(* Logix 5000 project; controller TFF vendor 1 type 14 code 107 rev 33.11; software revision 33.04; part 34 of 38 *)
(* tags used below, declared in another part *)
   Address : DINT;   // Temp Address
   Index : DINT;   // Index
   Index2 : DINT;   // Index
   _150S1 : ALIAS FOR DigitalOutput[0];
   AC008 : ALIAS FOR DigitalOutput[7];
   AlarmControl : AlarmControl;   // Alarm Control
   ALM001 : ALIAS FOR DigitalOutput[2];
   ALM002 : ALIAS FOR DigitalOutput[17];
   AnalogOutput : AnalogOutput[25];   // Analog Output Array
   AO1 : ALIAS FOR AnalogOutput[8];
   AO2 : ALIAS FOR AnalogOutput[9];
   AO3 : ALIAS FOR AnalogOutput[10];
   AO4 : ALIAS FOR AnalogOutput[11];
   AP008 : ALIAS FOR DigitalOutput[14];
   BAN001P : ALIAS FOR DigitalOutput[4];
   BAN001S : ALIAS FOR DigitalOutput[3];
   BAN002P : ALIAS FOR DigitalOutput[6];
   BAN002S : ALIAS FOR DigitalOutput[5];
   DigitalOutput : BOOL[256];   // Digital Output Array these bits are sent to output cards.
   DO1 : ALIAS FOR DigitalOutput[80];
   DO2 : ALIAS FOR DigitalOutput[81];
   DO3 : ALIAS FOR DigitalOutput[82];
   DO4 : ALIAS FOR DigitalOutput[83];
   DO5 : ALIAS FOR DigitalOutput[84];
   DO6 : ALIAS FOR DigitalOutput[85];
   DO7 : ALIAS FOR DigitalOutput[86];
   FlowPath : FlowPath[64];   // Flow Path Array
   IBA001 : ALIAS FOR DigitalOutput[25];
   MIX101ON : ALIAS FOR DigitalOutput[16];
   Mixer : Mixer;   // Mixer config. structure
   PCV101 : ALIAS FOR AnalogPoint[3];
   PCV101_AO : ALIAS FOR AnalogOutput[3];
   PCV201 : ALIAS FOR AnalogPoint[4];
   PCV201_AO : ALIAS FOR AnalogOutput[4];
   POWERON : ALIAS FOR DigitalOutput[1];
   PTA001 : ALIAS FOR DigitalOutput[21];
   PTA101 : ALIAS FOR DigitalOutput[22];
   PTA201 : ALIAS FOR DigitalOutput[23];
   PTA401 : ALIAS FOR DigitalOutput[24];
   PTA601 : ALIAS FOR DigitalOutput[26];
   Rack_Murr_Node0_Smart : IO_Station;   // Status of Node 0 Smart
   Rack_Murr_Node1_TFF40 : IO_Station;   // Status of Node 1 TFF40
   Rack_Murr_Node1_TFF80 : IO_Station;   // Status of Node 1 TFF80
   SIC001 : ALIAS FOR Drive[1];
   SIC001_AO : ALIAS FOR AnalogOutput[0];
   SIC001_DO : ALIAS FOR DigitalOutput[8];
   SIC002 : ALIAS FOR Drive[2];
   SIC002_AO : ALIAS FOR AnalogOutput[1];
   SIC002_DO : ALIAS FOR DigitalOutput[9];
   SIC003_AO : ALIAS FOR AnalogOutput[2];
   SIC003_DO : ALIAS FOR DigitalOutput[15];
   SIC004 : ALIAS FOR Drive[3];
   SIC004_AO : ALIAS FOR AnalogOutput[5];
   SysControl : SysControl;   // General system status and command
   Tank : TankManagement;   // Tank Management
   TCU101 : ALIAS FOR AnalogPoint[18];
   TCU101_AO : ALIAS FOR AnalogOutput[6];
   TCU101ON : ALIAS FOR DigitalOutput[20];
   ThisSystem : SystemType;
   TNK101 : ALIAS FOR DigitalOutput[18];
   TNK102 : ALIAS FOR DigitalOutput[19];
   TNK103 : ALIAS FOR DigitalOutput[27];
   Valve : Valve[100];   // Valve Array
   ValveControl : ValveControl;   // Valve Control
   XV001 : ALIAS FOR Valve[0];
   XV002 : ALIAS FOR Valve[1];
   XV003 : ALIAS FOR Valve[2];
   XV004 : ALIAS FOR Valve[3];
   XV005 : ALIAS FOR Valve[4];
   XV006 : ALIAS FOR Valve[5];
   XV007 : ALIAS FOR Valve[6];
   XV101 : ALIAS FOR Valve[7];
   XV102 : ALIAS FOR Valve[8];
   XV201 : ALIAS FOR Valve[15];
   XV202 : ALIAS FOR Valve[16];
   XV401 : ALIAS FOR Valve[9];
   XV402 : ALIAS FOR Valve[10];
   XV403 : ALIAS FOR Valve[11];
   XV404 : ALIAS FOR Valve[12];
   XV405 : ALIAS FOR Valve[13];
   XV406 : ALIAS FOR Valve[14];
   XV701 : ALIAS FOR Valve[17];
   XV702 : ALIAS FOR Valve[18];
   XV703 : ALIAS FOR Valve[19];
   XV704 : ALIAS FOR Valve[20];
   Y500A : ALIAS FOR DigitalOutput[10];
   Y500B : ALIAS FOR DigitalOutput[11];
   Y501A : ALIAS FOR DigitalOutput[12];
   Y501B : ALIAS FOR DigitalOutput[13];
(* Process, continued *)

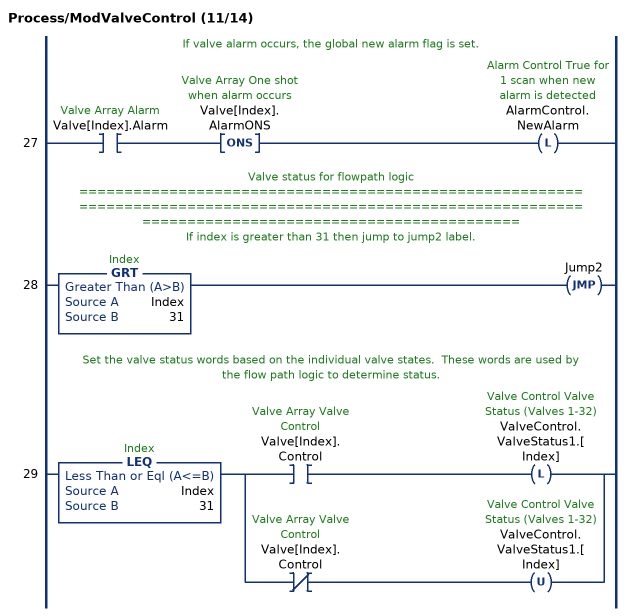
   [picture p422: Process/ModValveControl rungs 27-29]
   // If valve alarm occurs, the global new alarm flag is set.
   27: XIC(Valve[Index].Alarm)ONS(Valve[Index].AlarmONS)OTL(AlarmControl.NewAlarm);
   // Valve status for flowpath logic
   // ==========================================================================================================================================================
   // If index is greater than 31 then jump to jump2 label.
   28: GRT(Index,31)JMP(Jump2);
   // Set the valve status words based on the individual valve states.  These words are used by the flow path logic to determine status.
   29: LEQ(Index,31)[XIC(Valve[Index].Control) OTL(ValveControl.ValveStatus1.[Index]) ,XIO(Valve[Index].Control) OTU(ValveControl.ValveStatus1.[Index]) ];
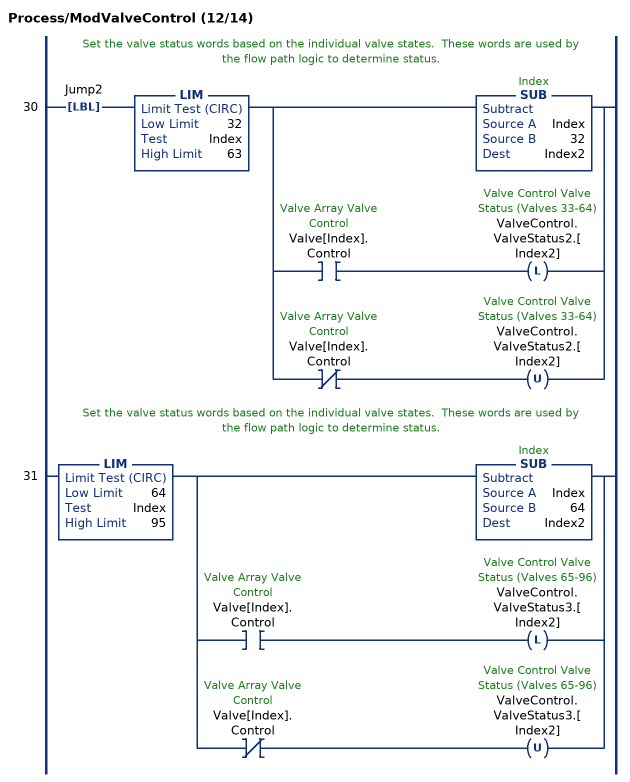
   // Set the valve status words based on the individual valve states.  These words are used by the flow path logic to determine status.
   30: LBL(Jump2)LIM(32,Index,63)[SUB(Index,32,Index2) ,XIC(Valve[Index].Control) OTL(ValveControl.ValveStatus2.[Index2]) ,XIO(Valve[Index].Control) OTU(ValveControl.ValveStatus2.[Index2]) ];
   // Set the valve status words based on the individual valve states.  These words are used by the flow path logic to determine status.
   31: LIM(64,Index,95)[SUB(Index,64,Index2) ,XIC(Valve[Index].Control) OTL(ValveControl.ValveStatus3.[Index2]) ,XIO(Valve[Index].Control) OTU(ValveControl.ValveStatus3.[Index2]) ];
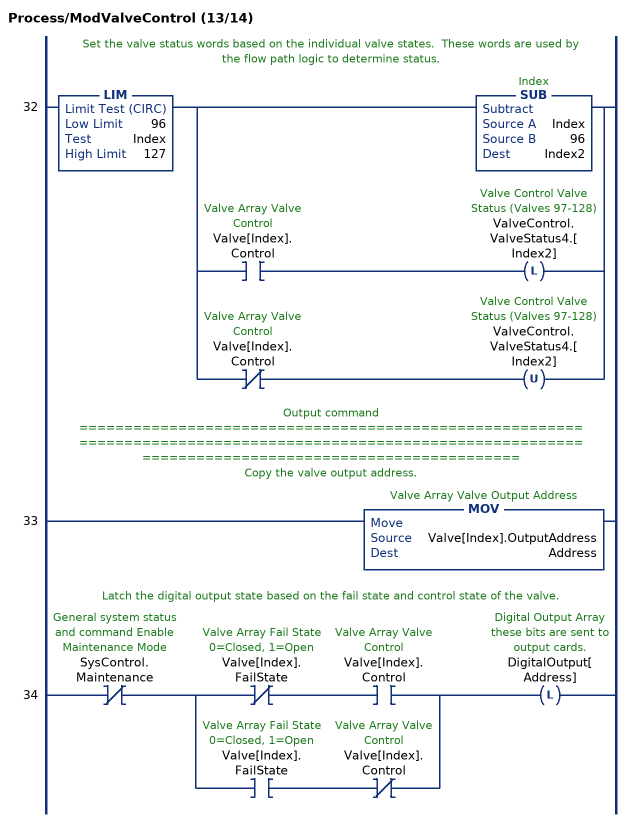
   // Set the valve status words based on the individual valve states.  These words are used by the flow path logic to determine status.
   32: LIM(96,Index,127)[SUB(Index,96,Index2) ,XIC(Valve[Index].Control) OTL(ValveControl.ValveStatus4.[Index2]) ,XIO(Valve[Index].Control) OTU(ValveControl.ValveStatus4.[Index2]) ];
   // Output command
   // ==========================================================================================================================================================
   // Copy the valve output address.
   33: MOV(Valve[Index].OutputAddress,Address);
   // Latch the digital output state based on the fail state and control state of the valve.
   34: XIO(SysControl.Maintenance)[XIO(Valve[Index].FailState) XIC(Valve[Index].Control) ,XIC(Valve[Index].FailState) XIO(Valve[Index].Control) ]OTL(DigitalOutput[Address]);
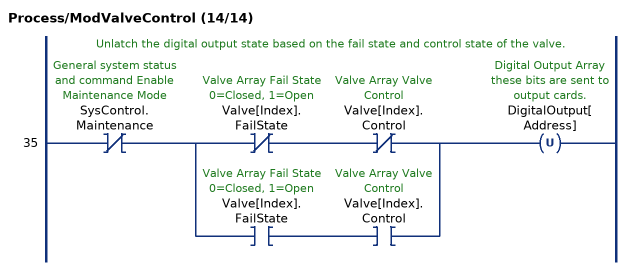
   // Unlatch the digital output state based on the fail state and control state of the valve.
   35: XIO(SysControl.Maintenance)[XIO(Valve[Index].FailState) XIO(Valve[Index].Control) ,XIC(Valve[Index].FailState) XIC(Valve[Index].Control) ]OTU(DigitalOutput[Address]);
END_ROUTINE

ROUTINE OutputAnalogPoint   (* ladder *)
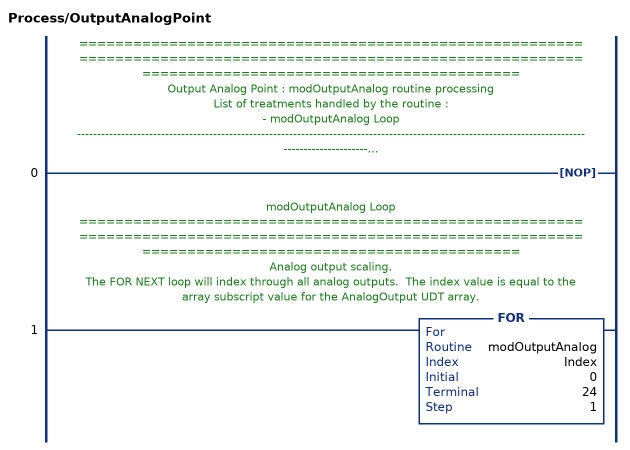
   // ==========================================================================================================================================================
   //                                                                                                             Output Analog Point : modOutputAnalog routine processing
   //                                                     List of treatments handled by the routine :
   //                                                          - modOutputAnalog Loop
   //                                                     -----------------------------------------------------------------------------------------------------------------------------------------------------
   //                                                     History
   // 		2019-DEC-24 - Merck - Q. Spindler - Initial version for Candidate Release 1.00.00.00.a
   // ==========================================================================================================================================================
   0: NOP();
   // modOutputAnalog Loop
   // ==========================================================================================================================================================
   // Analog output scaling.
   // The FOR NEXT loop will index through all analog outputs.  The index value is equal to the array subscript value for the AnalogOutput UDT array.
   1: FOR(modOutputAnalog,Index,0,24,1);
END_ROUTINE

ROUTINE OutputAnalogRaw   (* ladder *)
// Output Routine
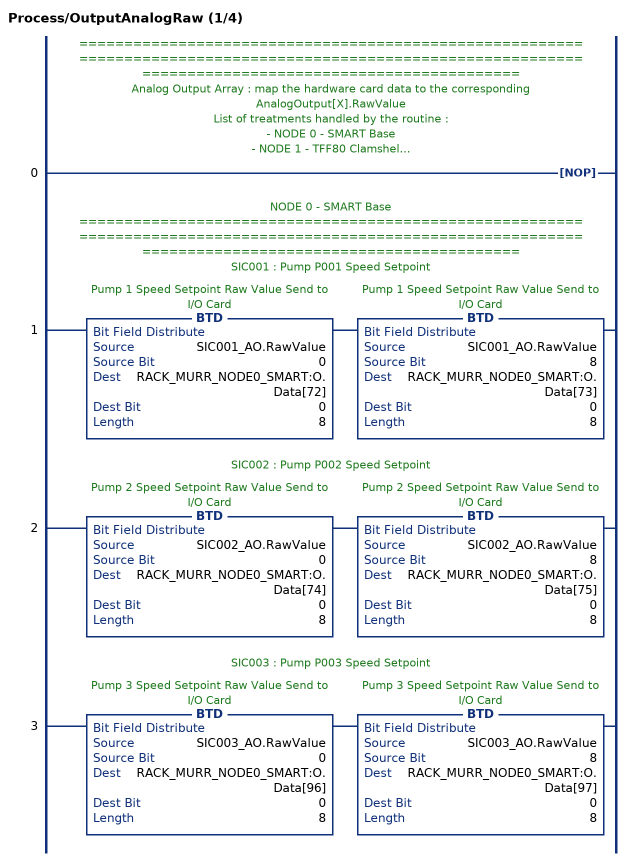
   // ==========================================================================================================================================================
   //                                                                                    Analog Output Array : map the hardware card data to the corresponding AnalogOutput[X].RawValue
   //                                                     List of treatments handled by the routine :
   //                                                    - NODE 0 - SMART Base
   //                                                         - NODE 1 - TFF80 Clamshell
   //                                                         - NODE 1 - TFF40 Clamshell
   //                                                         - NODE 1 - TFF20 Clamshell
   //                                                     -----------------------------------------------------------------------------------------------------------------------------------------------------
   //                                                     History
   // 		2019-DEC-24 - Merck - Q. Spindler - Initial version for Candidate Release 1.00.00.00.a
   // ==========================================================================================================================================================
   0: NOP();
   // NODE 0 - SMART Base
   // ==========================================================================================================================================================
   // SIC001 : Pump P001 Speed Setpoint
   1: BTD(SIC001_AO.RawValue,0,RACK_MURR_NODE0_SMART:O.Data[72],0,8)BTD(SIC001_AO.RawValue,8,RACK_MURR_NODE0_SMART:O.Data[73],0,8);
   // SIC002 : Pump P002 Speed Setpoint
   2: BTD(SIC002_AO.RawValue,0,RACK_MURR_NODE0_SMART:O.Data[74],0,8)BTD(SIC002_AO.RawValue,8,RACK_MURR_NODE0_SMART:O.Data[75],0,8);
   // SIC003 : Pump P003 Speed Setpoint
   3: BTD(SIC003_AO.RawValue,0,RACK_MURR_NODE0_SMART:O.Data[96],0,8)BTD(SIC003_AO.RawValue,8,RACK_MURR_NODE0_SMART:O.Data[97],0,8);
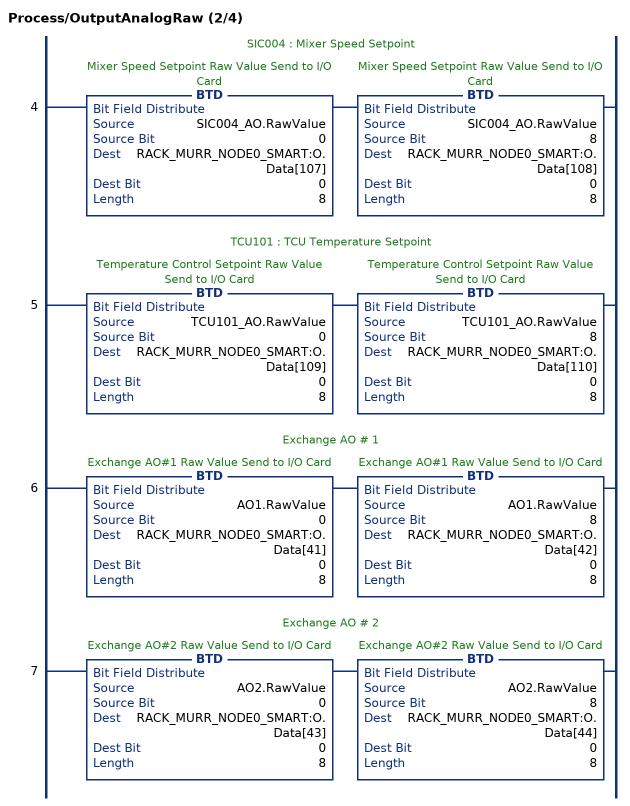
   // SIC004 : Mixer Speed Setpoint
   4: BTD(SIC004_AO.RawValue,0,RACK_MURR_NODE0_SMART:O.Data[107],0,8)BTD(SIC004_AO.RawValue,8,RACK_MURR_NODE0_SMART:O.Data[108],0,8);
   // TCU101 : TCU Temperature Setpoint
   5: BTD(TCU101_AO.RawValue,0,RACK_MURR_NODE0_SMART:O.Data[109],0,8)BTD(TCU101_AO.RawValue,8,RACK_MURR_NODE0_SMART:O.Data[110],0,8);
   // Exchange AO # 1
   6: BTD(AO1.RawValue,0,RACK_MURR_NODE0_SMART:O.Data[41],0,8)BTD(AO1.RawValue,8,RACK_MURR_NODE0_SMART:O.Data[42],0,8);
   // Exchange AO # 2
   7: BTD(AO2.RawValue,0,RACK_MURR_NODE0_SMART:O.Data[43],0,8)BTD(AO2.RawValue,8,RACK_MURR_NODE0_SMART:O.Data[44],0,8);
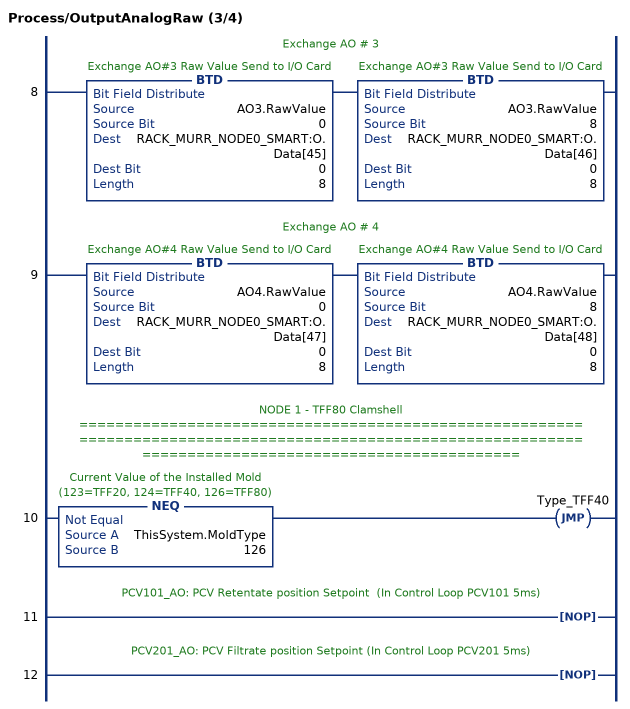
   // Exchange AO # 3
   8: BTD(AO3.RawValue,0,RACK_MURR_NODE0_SMART:O.Data[45],0,8)BTD(AO3.RawValue,8,RACK_MURR_NODE0_SMART:O.Data[46],0,8);
   // Exchange AO # 4
   9: BTD(AO4.RawValue,0,RACK_MURR_NODE0_SMART:O.Data[47],0,8)BTD(AO4.RawValue,8,RACK_MURR_NODE0_SMART:O.Data[48],0,8);
   // NODE 1 - TFF80 Clamshell
   // ==========================================================================================================================================================
   10: NEQ(ThisSystem.MoldType,126)JMP(Type_TFF40);
   // PCV101_AO: PCV Retentate position Setpoint  (In Control Loop PCV101 5ms)
   11: NOP();
   // PCV201_AO: PCV Filtrate position Setpoint (In Control Loop PCV201 5ms)
   12: NOP();
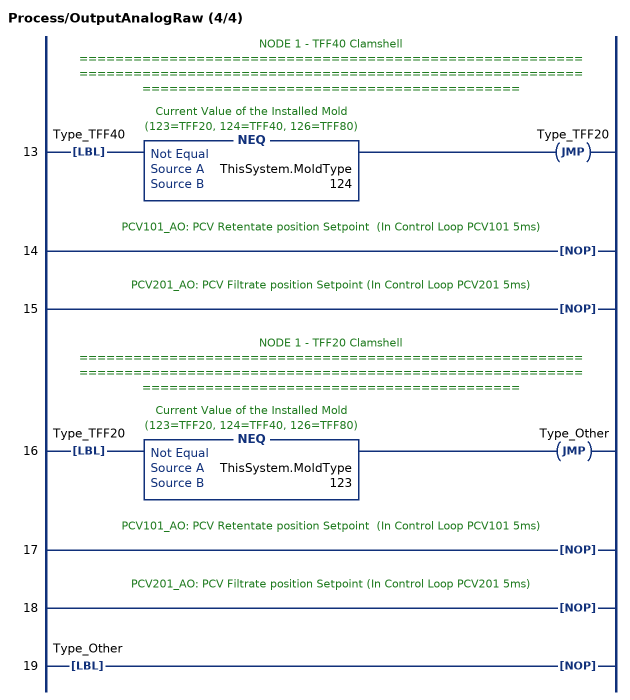
   // NODE 1 - TFF40 Clamshell
   // ==========================================================================================================================================================
   13: LBL(Type_TFF40)NEQ(ThisSystem.MoldType,124)JMP(Type_TFF20);
   // PCV101_AO: PCV Retentate position Setpoint  (In Control Loop PCV101 5ms)
   14: NOP();
   // PCV201_AO: PCV Filtrate position Setpoint (In Control Loop PCV201 5ms)
   15: NOP();
   // NODE 1 - TFF20 Clamshell
   // ==========================================================================================================================================================
   16: LBL(Type_TFF20)NEQ(ThisSystem.MoldType,123)JMP(Type_Other);
   // PCV101_AO: PCV Retentate position Setpoint  (In Control Loop PCV101 5ms)
   17: NOP();
   // PCV201_AO: PCV Filtrate position Setpoint (In Control Loop PCV201 5ms)
   18: NOP();
   19: LBL(Type_Other)NOP();
END_ROUTINE

ROUTINE OutputDigitalRaw   (* ladder *)
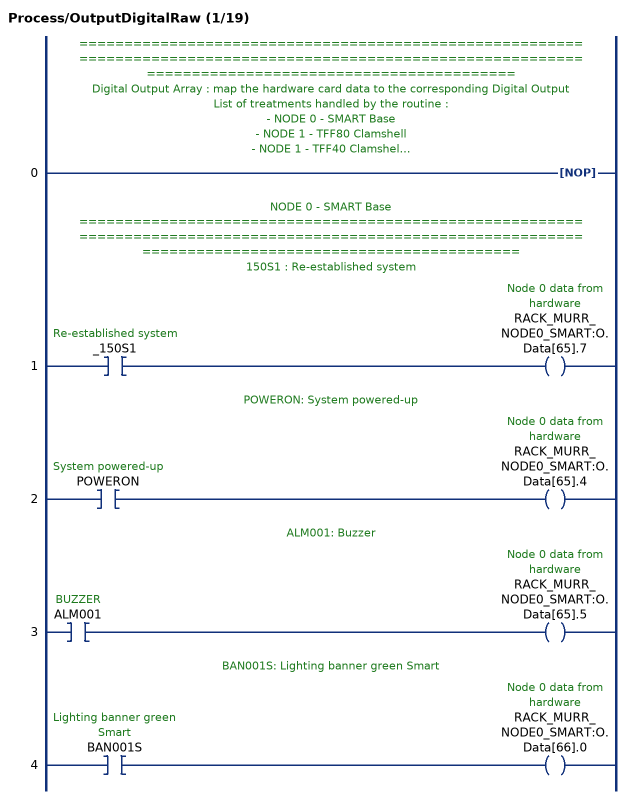
   // =========================================================================================================================================================
   //                                                                                          Digital Output Array : map the hardware card data to the corresponding Digital Output
   //                                                     List of treatments handled by the routine :
   //                                                    - NODE 0 - SMART Base
   //                                                         - NODE 1 - TFF80 Clamshell
   //                                                         - NODE 1 - TFF40 Clamshell
   //                                                         - NODE 1 - TFF20 Clamshell
   //                                                     -----------------------------------------------------------------------------------------------------------------------------------------------------
   //                                                     History
   // 		2019-DEC-24 - Merck - Q. Spindler - Initial version for Candidate Release 1.00.00.00.a
   // 		2020-MAR-30 - Merck - Q. Spindler - Initial version for Candidate Release 1.00.00.00.b
   //                                           - Change IO mapping for External DOs and PTA101 and PTA401
   // - Add TNK103 : Feed Tank Weight Zero
   // ==========================================================================================================================================================
   0: NOP();
   // NODE 0 - SMART Base
   // ==========================================================================================================================================================
   // 150S1 : Re-established system
   1: XIC(_150S1)OTE(RACK_MURR_NODE0_SMART:O.Data[65].7);
   // POWERON: System powered-up
   2: XIC(POWERON)OTE(RACK_MURR_NODE0_SMART:O.Data[65].4);
   // ALM001: Buzzer
   3: XIC(ALM001)OTE(RACK_MURR_NODE0_SMART:O.Data[65].5);
   // BAN001S: Lighting banner green Smart
   4: XIC(BAN001S)OTE(RACK_MURR_NODE0_SMART:O.Data[66].0);
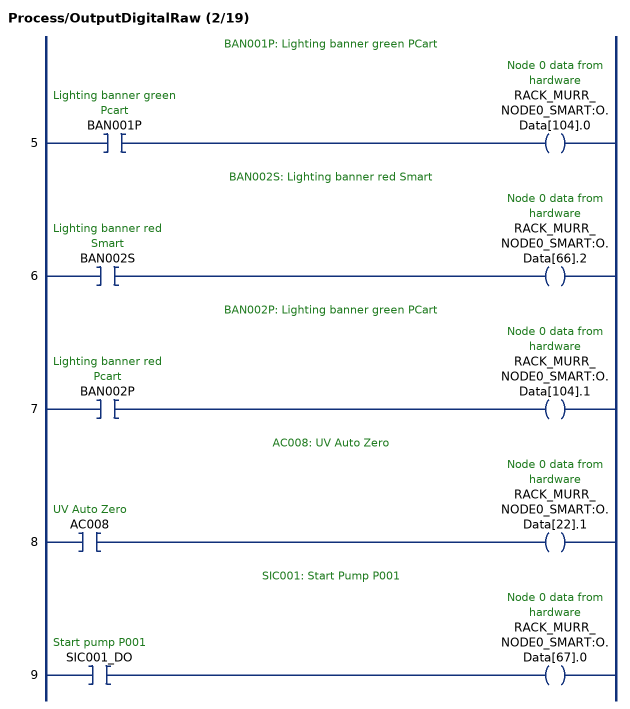
   // BAN001P: Lighting banner green PCart
   5: XIC(BAN001P)OTE(RACK_MURR_NODE0_SMART:O.Data[104].0);
   // BAN002S: Lighting banner red Smart
   6: XIC(BAN002S)OTE(RACK_MURR_NODE0_SMART:O.Data[66].2);
   // BAN002P: Lighting banner green PCart
   7: XIC(BAN002P)OTE(RACK_MURR_NODE0_SMART:O.Data[104].1);
   // AC008: UV Auto Zero
   8: XIC(AC008)OTE(RACK_MURR_NODE0_SMART:O.Data[22].1);
   // SIC001: Start Pump P001
   9: XIC(SIC001_DO)OTE(RACK_MURR_NODE0_SMART:O.Data[67].0);
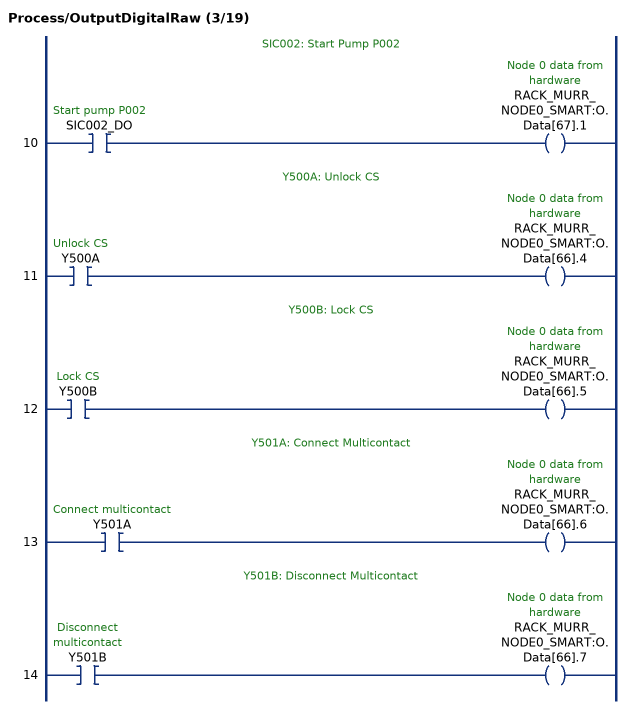
   // SIC002: Start Pump P002
   10: XIC(SIC002_DO)OTE(RACK_MURR_NODE0_SMART:O.Data[67].1);
   // Y500A: Unlock CS
   11: XIC(Y500A)OTE(RACK_MURR_NODE0_SMART:O.Data[66].4);
   // Y500B: Lock CS
   12: XIC(Y500B)OTE(RACK_MURR_NODE0_SMART:O.Data[66].5);
   // Y501A: Connect Multicontact
   13: XIC(Y501A)OTE(RACK_MURR_NODE0_SMART:O.Data[66].6);
   // Y501B: Disconnect Multicontact
   14: XIC(Y501B)OTE(RACK_MURR_NODE0_SMART:O.Data[66].7);
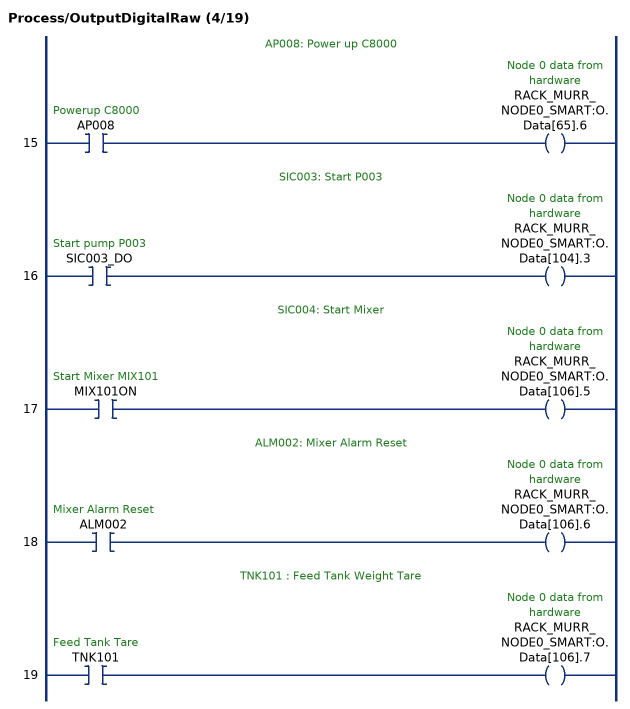
   // AP008: Power up C8000
   15: XIC(AP008)OTE(RACK_MURR_NODE0_SMART:O.Data[65].6);
   // SIC003: Start P003
   16: XIC(SIC003_DO)OTE(RACK_MURR_NODE0_SMART:O.Data[104].3);
   // SIC004: Start Mixer
   17: XIC(MIX101ON)OTE(RACK_MURR_NODE0_SMART:O.Data[106].5);
   // ALM002: Mixer Alarm Reset
   18: XIC(ALM002)OTE(RACK_MURR_NODE0_SMART:O.Data[106].6);
   // TNK101 : Feed Tank Weight Tare
   19: XIC(TNK101)OTE(RACK_MURR_NODE0_SMART:O.Data[106].7);
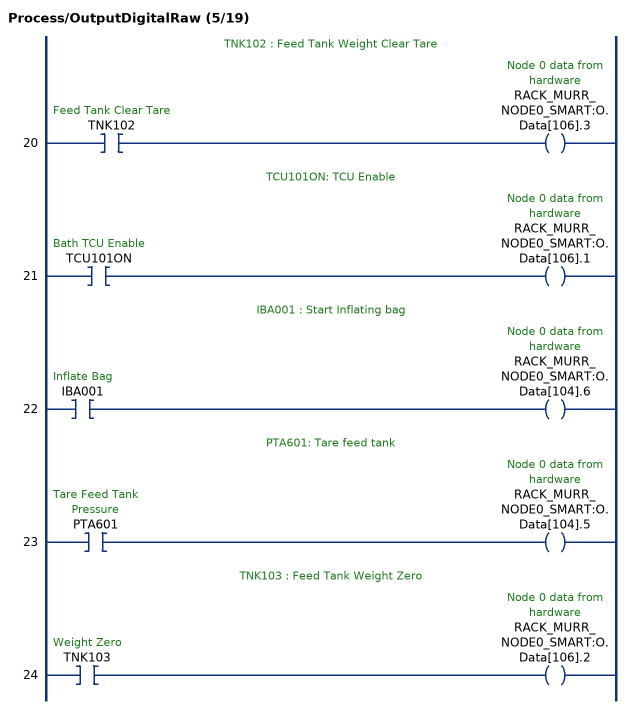
   // TNK102 : Feed Tank Weight Clear Tare
   20: XIC(TNK102)OTE(RACK_MURR_NODE0_SMART:O.Data[106].3);
   // TCU101ON: TCU Enable
   21: XIC(TCU101ON)OTE(RACK_MURR_NODE0_SMART:O.Data[106].1);
   // IBA001 : Start Inflating bag
   22: XIC(IBA001)OTE(RACK_MURR_NODE0_SMART:O.Data[104].6);
   // PTA601: Tare feed tank
   23: XIC(PTA601)OTE(RACK_MURR_NODE0_SMART:O.Data[104].5);
   // TNK103 : Feed Tank Weight Zero
   24: XIC(TNK103)OTE(RACK_MURR_NODE0_SMART:O.Data[106].2);
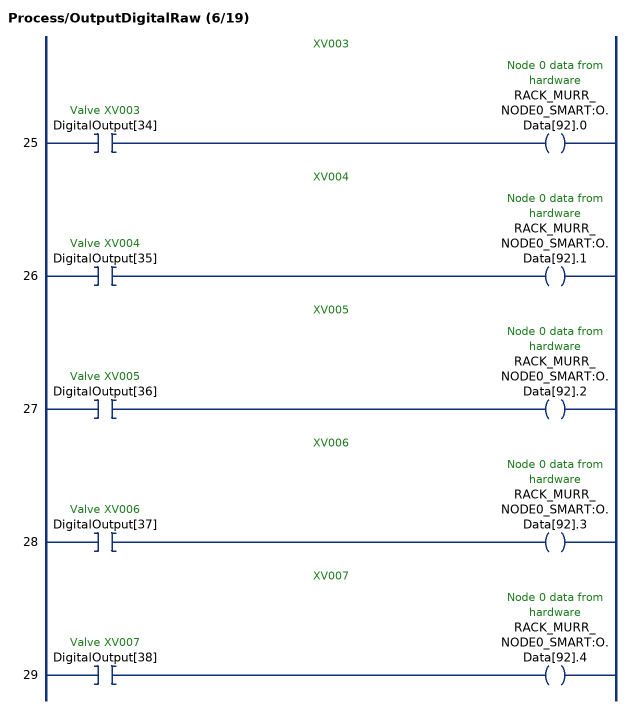
   // XV003
   25: XIC(DigitalOutput[34])OTE(RACK_MURR_NODE0_SMART:O.Data[92].0);
   // XV004
   26: XIC(DigitalOutput[35])OTE(RACK_MURR_NODE0_SMART:O.Data[92].1);
   // XV005
   27: XIC(DigitalOutput[36])OTE(RACK_MURR_NODE0_SMART:O.Data[92].2);
   // XV006
   28: XIC(DigitalOutput[37])OTE(RACK_MURR_NODE0_SMART:O.Data[92].3);
   // XV007
   29: XIC(DigitalOutput[38])OTE(RACK_MURR_NODE0_SMART:O.Data[92].4);
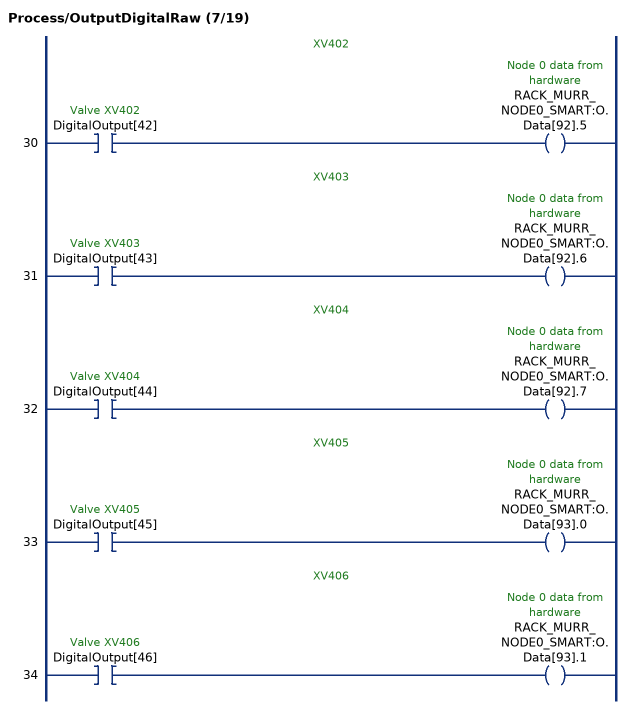
   // XV402
   30: XIC(DigitalOutput[42])OTE(RACK_MURR_NODE0_SMART:O.Data[92].5);
   // XV403
   31: XIC(DigitalOutput[43])OTE(RACK_MURR_NODE0_SMART:O.Data[92].6);
   // XV404
   32: XIC(DigitalOutput[44])OTE(RACK_MURR_NODE0_SMART:O.Data[92].7);
   // XV405
   33: XIC(DigitalOutput[45])OTE(RACK_MURR_NODE0_SMART:O.Data[93].0);
   // XV406
   34: XIC(DigitalOutput[46])OTE(RACK_MURR_NODE0_SMART:O.Data[93].1);
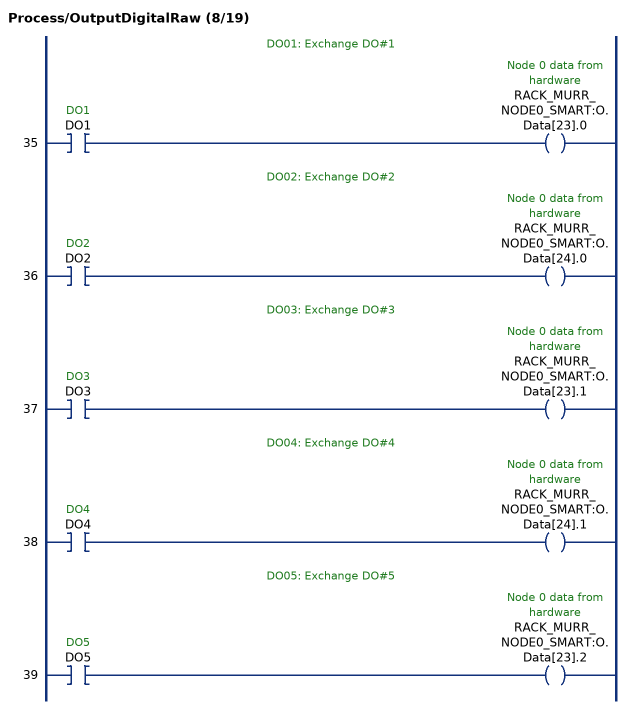
   // DO01: Exchange DO#1
   35: XIC(DO1)OTE(RACK_MURR_NODE0_SMART:O.Data[23].0);
   // DO02: Exchange DO#2
   36: XIC(DO2)OTE(RACK_MURR_NODE0_SMART:O.Data[24].0);
   // DO03: Exchange DO#3
   37: XIC(DO3)OTE(RACK_MURR_NODE0_SMART:O.Data[23].1);
   // DO04: Exchange DO#4
   38: XIC(DO4)OTE(RACK_MURR_NODE0_SMART:O.Data[24].1);
   // DO05: Exchange DO#5
   39: XIC(DO5)OTE(RACK_MURR_NODE0_SMART:O.Data[23].2);
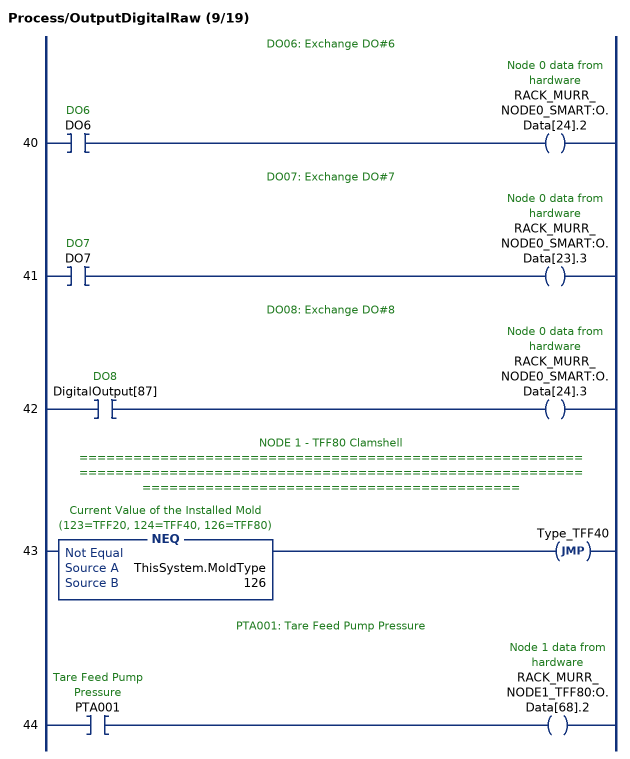
   // DO06: Exchange DO#6
   40: XIC(DO6)OTE(RACK_MURR_NODE0_SMART:O.Data[24].2);
   // DO07: Exchange DO#7
   41: XIC(DO7)OTE(RACK_MURR_NODE0_SMART:O.Data[23].3);
   // DO08: Exchange DO#8
   42: XIC(DigitalOutput[87])OTE(RACK_MURR_NODE0_SMART:O.Data[24].3);
   // NODE 1 - TFF80 Clamshell
   // ==========================================================================================================================================================
   43: NEQ(ThisSystem.MoldType,126)JMP(Type_TFF40);
   // PTA001: Tare Feed Pump Pressure
   44: XIC(PTA001)OTE(RACK_MURR_NODE1_TFF80:O.Data[68].2);
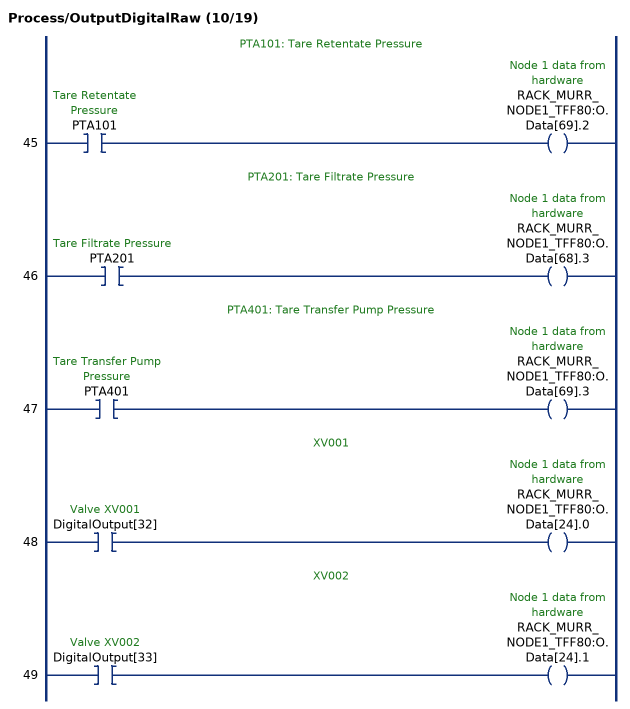
   // PTA101: Tare Retentate Pressure
   45: XIC(PTA101)OTE(RACK_MURR_NODE1_TFF80:O.Data[69].2);
   // PTA201: Tare Filtrate Pressure
   46: XIC(PTA201)OTE(RACK_MURR_NODE1_TFF80:O.Data[68].3);
   // PTA401: Tare Transfer Pump Pressure
   47: XIC(PTA401)OTE(RACK_MURR_NODE1_TFF80:O.Data[69].3);
   // XV001
   48: XIC(DigitalOutput[32])OTE(RACK_MURR_NODE1_TFF80:O.Data[24].0);
   // XV002
   49: XIC(DigitalOutput[33])OTE(RACK_MURR_NODE1_TFF80:O.Data[24].1);
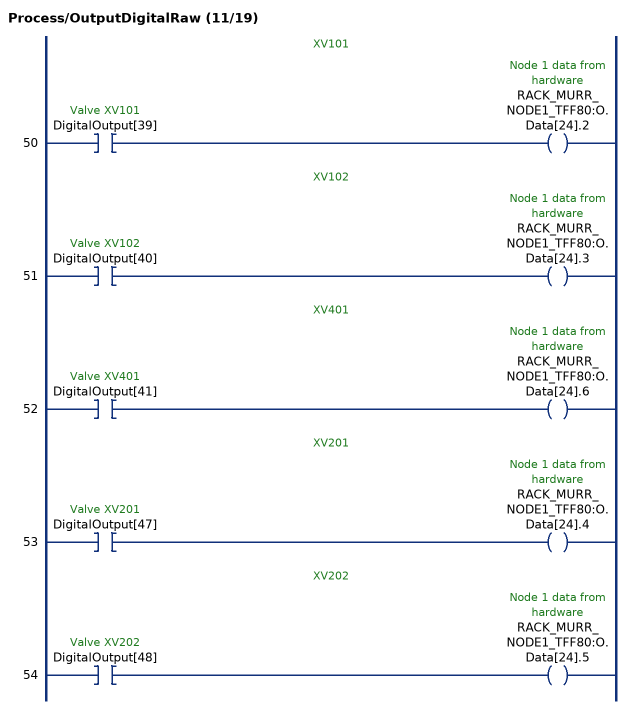
   // XV101
   50: XIC(DigitalOutput[39])OTE(RACK_MURR_NODE1_TFF80:O.Data[24].2);
   // XV102
   51: XIC(DigitalOutput[40])OTE(RACK_MURR_NODE1_TFF80:O.Data[24].3);
   // XV401
   52: XIC(DigitalOutput[41])OTE(RACK_MURR_NODE1_TFF80:O.Data[24].6);
   // XV201
   53: XIC(DigitalOutput[47])OTE(RACK_MURR_NODE1_TFF80:O.Data[24].4);
   // XV202
   54: XIC(DigitalOutput[48])OTE(RACK_MURR_NODE1_TFF80:O.Data[24].5);
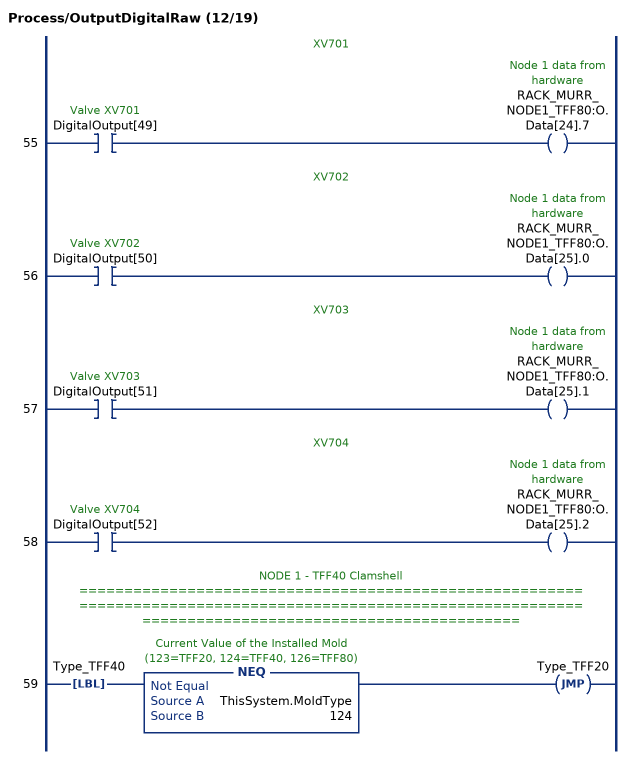
   // XV701
   55: XIC(DigitalOutput[49])OTE(RACK_MURR_NODE1_TFF80:O.Data[24].7);
   // XV702
   56: XIC(DigitalOutput[50])OTE(RACK_MURR_NODE1_TFF80:O.Data[25].0);
   // XV703
   57: XIC(DigitalOutput[51])OTE(RACK_MURR_NODE1_TFF80:O.Data[25].1);
   // XV704
   58: XIC(DigitalOutput[52])OTE(RACK_MURR_NODE1_TFF80:O.Data[25].2);
   // NODE 1 - TFF40 Clamshell
   // ==========================================================================================================================================================
   59: LBL(Type_TFF40)NEQ(ThisSystem.MoldType,124)JMP(Type_TFF20);
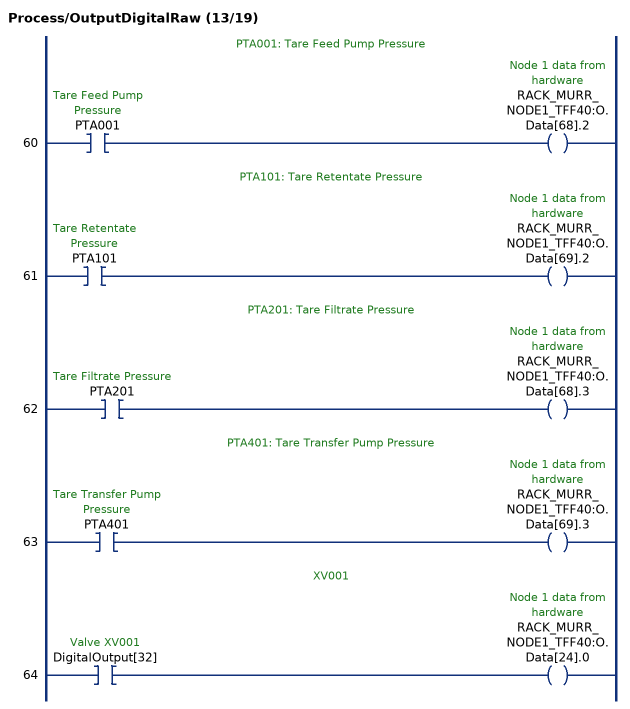
   // PTA001: Tare Feed Pump Pressure
   60: XIC(PTA001)OTE(RACK_MURR_NODE1_TFF40:O.Data[68].2);
   // PTA101: Tare Retentate Pressure
   61: XIC(PTA101)OTE(RACK_MURR_NODE1_TFF40:O.Data[69].2);
   // PTA201: Tare Filtrate Pressure
   62: XIC(PTA201)OTE(RACK_MURR_NODE1_TFF40:O.Data[68].3);
   // PTA401: Tare Transfer Pump Pressure
   63: XIC(PTA401)OTE(RACK_MURR_NODE1_TFF40:O.Data[69].3);
   // XV001
   64: XIC(DigitalOutput[32])OTE(RACK_MURR_NODE1_TFF40:O.Data[24].0);
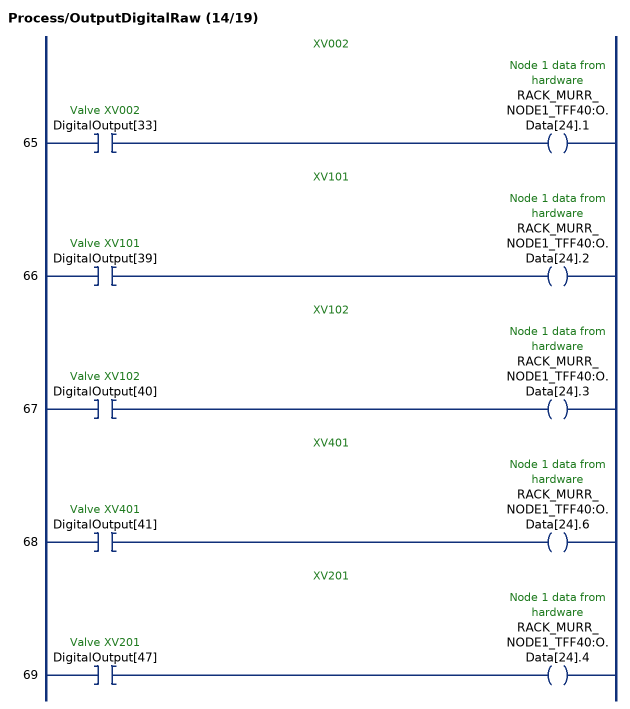
   // XV002
   65: XIC(DigitalOutput[33])OTE(RACK_MURR_NODE1_TFF40:O.Data[24].1);
   // XV101
   66: XIC(DigitalOutput[39])OTE(RACK_MURR_NODE1_TFF40:O.Data[24].2);
   // XV102
   67: XIC(DigitalOutput[40])OTE(RACK_MURR_NODE1_TFF40:O.Data[24].3);
   // XV401
   68: XIC(DigitalOutput[41])OTE(RACK_MURR_NODE1_TFF40:O.Data[24].6);
   // XV201
   69: XIC(DigitalOutput[47])OTE(RACK_MURR_NODE1_TFF40:O.Data[24].4);
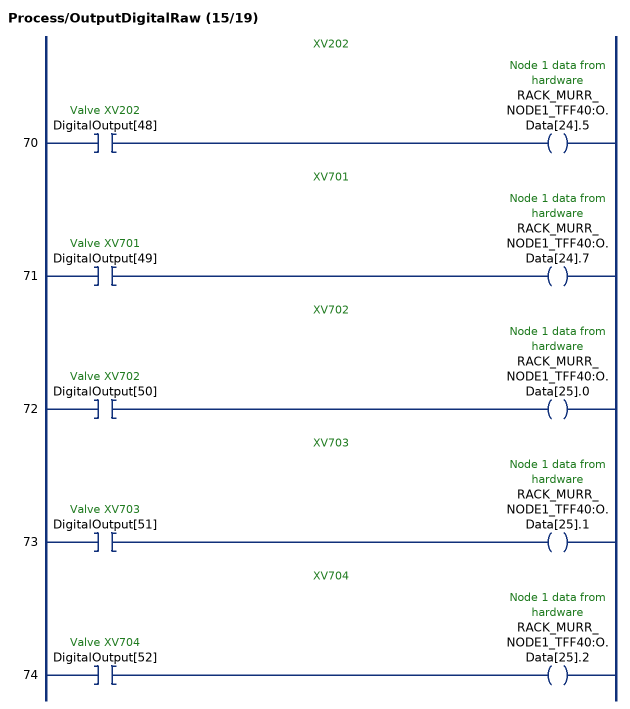
   // XV202
   70: XIC(DigitalOutput[48])OTE(RACK_MURR_NODE1_TFF40:O.Data[24].5);
   // XV701
   71: XIC(DigitalOutput[49])OTE(RACK_MURR_NODE1_TFF40:O.Data[24].7);
   // XV702
   72: XIC(DigitalOutput[50])OTE(RACK_MURR_NODE1_TFF40:O.Data[25].0);
   // XV703
   73: XIC(DigitalOutput[51])OTE(RACK_MURR_NODE1_TFF40:O.Data[25].1);
   // XV704
   74: XIC(DigitalOutput[52])OTE(RACK_MURR_NODE1_TFF40:O.Data[25].2);
